Staubli VAL3: start.pgx

program start()
// Isma structure adapted to Level 2; taught joints, bounded cycles and shared IO modes.
  local num poseIndex
  local point approachPose
  local point placePose
  local point pistonApproach
begin
  // ============================================================
  // LEVEL 2: ALIMENTAR, MONTAR Y COLOCAR CUATRO CONJUNTOS
  // ============================================================
  // Adaptacion Level 2 de la estructura de Isma; originales preservados.
  // Lab2B (Level 1) y Lab2B_Level2 permanecen sin modificar.
  // Matriz VACIA y cuatro pistones cargados al comenzar.
  // simulation=true: sensores manuales, sin acceso a pines.
  // simulation=false: bIn2/14/15, bOut10 y pinza valve1.
  userPage()
  cls()
  putln("Lab2B_IsmaL2 - Four assemblies - empty matrix required")
  physicalRun = !simulation
  placedCount = 0
  partIndex = 0
  cycleStep = 0
  feederExtend = false
  ioReady = false

  // ============================================================
  // COMPROBAR ALTURAS DE MATRIZ SIN MOVER NI ACCIONAR SALIDAS
  // ============================================================
  // Parejas 0/1, 2/3, 4/5, 6/7: par=approach, impar=deposito.
  // J3 es un ANGULO, no una altura. Calculamos Z del TCP lateral.
  // Esto comprueba altura, no colisiones, alineacion o alcance del trayecto.
  for poseIndex = 0 to 3
    approachPose = jointToPoint(tLateral, world, jMatrix[2*poseIndex])
    placePose = jointToPoint(tLateral, world, jMatrix[2*poseIndex+1])
    putln("Matrix slot (0..3):")
    putln(poseIndex)
    putln("Approach Z (mm):")
    putln(approachPose.trsf.z)
    putln("Place Z (mm):")
    putln(placePose.trsf.z)
    if approachPose.trsf.z <= placePose.trsf.z
      putln("ERROR: approach is not above place; review this matrix pair")
      return
    endIf
  endFor

  // ============================================================
  // CUATRO RECOGIDAS REALES: IMG_3805, 3806, 3807, 3808
  // ============================================================
  // Impares = recogidas ensenadas; pares = aproximaciones calculadas.
  // Subir en Z de world conservando orientacion y configuracion del TCP.
  // El calculo termina antes de crear tareas o accionar el robot.
  if pistonLift <= 0
    putln("ERROR: pistonLift must be positive (mm)")
    return
  endIf
  for poseIndex = 0 to 3
    if jPistonPick[2*poseIndex+1].j1 == 0 and jPistonPick[2*poseIndex+1].j2 == 0 and jPistonPick[2*poseIndex+1].j3 == 0 and jPistonPick[2*poseIndex+1].j4 == 0 and jPistonPick[2*poseIndex+1].j5 == 0 and jPistonPick[2*poseIndex+1].j6 == 0
      putln("ERROR: teach piston pick joint; missing piston (0..3):")
      putln(poseIndex)
      return
    endIf
    pistonApproach = jointToPoint(tTip, world, jPistonPick[2*poseIndex+1])
    pistonApproach.trsf.z = pistonApproach.trsf.z + pistonLift
    if !pointToJoint(tTip, jPistonPick[2*poseIndex+1], pistonApproach, jPistonPick[2*poseIndex])
      putln("ERROR: no piston approach solution; piston (0..3):")
      putln(poseIndex)
      return
    endIf
    putln("Piston approach computed; piston (0..3):")
    putln(poseIndex)
    putln("World Z lift (mm):")
    putln(pistonLift)
  endFor

  // physicalIO solo escribe el ALIMENTADOR; nunca la pinza.
  if physicalRun
    taskCreate "physicalIO", 10, physicalIO()
    wait(ioReady == true)
    putln("PHYSICAL: real sensors and feeder enabled")
    open(tLateral)
  else
    putln("MANUAL SIMULATION: change sensor bools at the indicated steps")
    delay(tLateral.otime)
  endIf
  movej(jStart[0], tLateral, mNomSpeed)
  waitEndMove()

  // ============================================================
  // SOLO CUATRO CONJUNTOS; NO HAY QUINTA ALIMENTACION
  // ============================================================
  while placedCount < 4
    partIndex = placedCount
    putln("Assembly number (1..4):")
    putln(partIndex+1)
    call feedCylinder()
    call placeCylinder()
    call insertPiston()
    call placeInMatrix()
    // Contar tras soltar y terminar la retirada de la matriz.
    placedCount = placedCount + 1
    putln("Completed matrix slots:")
    putln(placedCount)
    // Volver a la postura inicial SOLO si falta otro conjunto.
    if placedCount < 4
      movej(jStart[0], tLateral, mNomSpeed)
      waitEndMove()
    endIf
  endWhile

  // La matriz llena finaliza aunque bIn2 siga detectando cilindros.
  feederExtend = false
  taskKill("physicalIO")
  if physicalRun
    io:bOut10 = false
  endIf
  ioReady = false
  cycleStep = 100
  putln("100 - Matrix full: 4/4. No further feeding or pickup.")
end
